Fanuc KAREL source: kt00403.KL

-- PROVISIONAL review KL for V770-1; original PC SHA256 26553de3f4d6d7f6d9013818d098ce96b3de3427f4c87bacff4e1eed68527ece
-- Incomplete behavior may be omitted. Consult companion uncertainty JSON. Do not deploy.
PROGRAM KT00403
%NOLOCKGROUP
VAR
  I1 : INTEGER
  OUT : BOOLEAN
-- UNRESOLVED_DECL Y2 type=002018
BEGIN
  -- UNRESOLVED_PC offsets 5-16; opcodes 2E,23
  -- UNRESOLVED_PC offsets 21-35; opcodes 2E,22,9D,33,B2
  -- UNRESOLVED_PC offsets 40-62; opcodes 21,22,9D,33,B1,5B,23
  -- UNRESOLVED_PC offsets 67-71; opcodes 7F
END KT00403
